(* IEC 61131-3 sources: repolevel_ST_code_completion/extract_code/重型运输系统/can/struct, 12 files *)

(* ---- Can_baseframe.st ---- *)
TYPE Can_baseframe :
STRUCT
	id		: UINT;
	data	: ARRAY[1..8] OF BYTE;
END_STRUCT
END_TYPE

(* ---- Can_BUS_8Inputs.st ---- *)
TYPE Can_BUS_8Inputs :          //输入缓存结构 EL2721-8Message_IN
STRUCT
	TxCounter			: UINT;
	RxCounter			: UINT;
	NoOfRxMessages 	 	: UINT;
	TransactionNumber	: UINT;
	RXMsg				: ARRAY[1..8] OF Can_Bus_RXMsg_Buff;
	CAN_State			: UINT;
	Align				: UINT;
	RX_Error_Cnt		: BYTE;
	TX_Error_Cnt		: BYTE;
END_STRUCT
END_TYPE

(* ---- Can_BUS_8Outputs.st ---- *)
TYPE Can_BUS_8Outputs :		//输出缓存结构 EL2721-8Message_OUT
STRUCT
	TxCounter		: UINT;
	RxCounter		: UINT;
	NoOfTxMessages 	: UINT;
	TXMsg			: ARRAY[1..8] OF Can_Bus_TXMsg_Buff;
	CAN_Control		: UINT;
END_STRUCT
END_TYPE

(* ---- Can_Bus_RXMsg_Buff.st ---- *)
TYPE Can_Bus_RXMsg_Buff:
STRUCT
	RxMsg_CobId		: UINT;
	RxMsg_Byte  	: ARRAY[1..8] OF BYTE;
END_STRUCT
END_TYPE

(* ---- Can_Bus_TXMsg_Buff.st ---- *)
TYPE Can_Bus_TXMsg_Buff :
STRUCT
	TxMsg_TransactionNumber		: UINT;
	TxMsg_CobId					: UINT;
	TxMsg_Byte  				: ARRAY[1..8] OF BYTE;
END_STRUCT
END_TYPE

(* ---- CmdPercentSet.st ---- *)
TYPE CmdPercentSet :
STRUCT
	extendPercent		:WORD;		//0-65535
	retractPercent		:WORD;		//0-65535
END_STRUCT
END_TYPE

(* ---- DeviceUnit.st ---- *)
TYPE DeviceUnit :
STRUCT

	sensor			:SensorInfo;		//传感器参数
	ctrl			:DevPid;			//pid等计算控制执行参数

	vector			:TargetDirect;		//指令运行方向 1-伸出 2-缩回 3-停止
	state			:DevStatus;			//设备状态 0-未知 1-运行 2-伸出到位 3-缩回到位 4-错误

	timeCounter		:INT;				//timeoutCounter超时计数器
	exeCounter		:INT;				//ExecuteCounter额外执行时间计数

	current			:ARRAY[1..2] OF WORD;	//电流mA	[i,j] -> 地轨挡板i的电流，j=1伸出电流，j=2缩回电流

END_STRUCT
END_TYPE

(* ---- DevStatus.st ---- *)
{attribute 'qualified_only'}
{attribute 'strict'}
TYPE DevStatus :
(
	unknown 	:= 0,

	runing		:= 1,

	extended	:= 2,

	retracted	:= 3,

	error		:= 4
);
END_TYPE

(* ---- SensorInfo.st ---- *)
TYPE SensorInfo :
STRUCT

	position	:REAL;	//实时位移
	speed		:REAL;	//实时速度

	//记录最大最小位移值
	retractVal	:REAL;	//缩回到位值
	extendVal	:REAL;	//伸出到位值

END_STRUCT
END_TYPE

(* ---- TargetDirect.st ---- *)
{attribute 'qualified_only'}
{attribute 'strict'}
TYPE TargetDirect :
(
	extend 	:= 1,	//伸出

	retract := 2,	//缩回

	stop	:= 3	//停止
);
END_TYPE

(* ---- UIMode.st ---- *)
TYPE UIMode :
STRUCT
	manualButtonSet			:BOOL;		//手动复位按钮模式
	usePID					:BOOL;		//使用pid
	autoEnable				:BOOL;		//自动使能
	manualPercentSet		:BOOL;		//手动设定比例量
	manualSetPid			:BOOL;		//手动调节pid参数，可通过pid测试界面设定目标位移值

	syncExt					:BOOL;		//同步伸
	syncRct					:BOOL;		//同步缩

	hydPowerOn				:BOOL;		//液压站开启 modbus 使用
	hydPowerOff				:BOOL;		//液压站关闭 modbus 使用
	hydPowerReset			:BOOL;
END_STRUCT
END_TYPE

(* ---- UIUnit.st ---- *)
TYPE UIUnit :
STRUCT
	//cmd
	pwrEnable			:BOOL;		//比例阀使能   power-enable
	pwrPercent			:REAL;		//比例阀百分比 power-percent 0-100

	//button
	btnExtend			:BOOL;
	btnRetract			:BOOL;
	btnStop				:BOOL;
	btnLast				:TargetDirect;	//上次动作方向

	//info display
	name				:STRING;	//挡板名
	wname				:WSTRING;	//山河命名
	hzname				:WSTRING;	//hua zhong ming ming
	postion				:REAL;		//位移值
	speed				:REAL;
	extendPercent		:REAL;		//伸出百分比 extend-percent

END_STRUCT
END_TYPE
